(* IEC 61131-3 sources: s7-to-codesys/src/POUs/S7Compat/F_S5RetOnDelay, 2 files *)

(* ---- F_S5RetOnDelay.decl.st ---- *)
// Назначение: SS T n — таймер S5 «задержка включения с памятью» (S_ODTS). Фронт RLO 0 → 1 запускает таймер
//             (идущий — перезапускает), время истекает независимо от RLO; Q = TRUE по истечении и держится
//             до сброса R (AWL_e.pdf §12.10, LAD §13.6). Возвращает Q после инструкции.
// Автор:      kr0nsch
// Версия:     1.2.0
// Документ:   docs/MAPPING_STL.md, правило s5.timebase
FUNCTION F_S5RetOnDelay : BOOL
VAR_IN_OUT
    stTimer : ST_S5Timer;   // таймер (GVL_S5Timers.aTimer[n])
END_VAR
VAR_INPUT
    xRlo : BOOL;            // RLO перед инструкцией
    wS5Time : WORD;         // заданное время S5TIME (ACCU1-L)
END_VAR

(* ---- F_S5RetOnDelay.impl.st ---- *)
stTimer.xQAtEnd := TRUE;
IF xRlo AND NOT stTimer.xRloStart THEN
    F_S5Start(stTimer := stTimer, wS5Time := wS5Time);
END_IF
stTimer.xRloStart := xRlo;
F_S5RetOnDelay := stTimer.xQ;
